(* IEC 61131-3 sources: kauha-loader-autonomy/plc/codesys/src/codesys_only, 3 files *)

(* ---- GVL_IO.st ---- *)
(* Hardware I/O of the 1:8 testbed safety PLC. Map each variable to its channel in
   the device's "I/O Mapping" tab (Raspberry Pi GPIOs device, or the I/O modules of
   your controller). Pin numbers are the testbed wiring in docs/scale/wiring.md.
   Inputs arrive through the 24 V opto-isolated input board (high = 24 V present). *)
VAR_GLOBAL
    (* inputs *)
    xEstopChainOk    : BOOL;   (* IN1  GPIO5:  safety relay K1 contact 33-34, TRUE = chain closed and K1 reset *)
    xRelayFeedbackOk : BOOL;   (* IN2  GPIO6:  K-DRIVE and K-IMPL NC mirror contacts in series, TRUE = both dropped *)
    stScannerIO      : ST_ScannerIO;
                               (* IN3  GPIO12: front_ossd_clear   IN4  GPIO13: rear_ossd_clear
                                  IN5  GPIO19: front_warn_clear   IN6  GPIO20: rear_warn_clear
                                  IN7  GPIO21: side_clear         IN8  GPIO26: under_clear
                                  scanners_ready: IN3..IN8 board "power good" (GPIO4) *)
    (* outputs *)
    xDriveEnable     : BOOL;   (* OUT1 GPIO23: coil of K-DRIVE (motor power and dynamic-brake changeover) *)
    xImplementEnable : BOOL;   (* OUT2 GPIO24: coil of K-IMPL (actuator power) *)
    xFs0, xFs1, xFs2, xFs3, xFs4, xFs5 : BOOL;
                               (* OUT3..OUT8 GPIO16, 17, 22, 27, 18, 14: field-set code bits 0..5 to the
                                  rated scanners' static control inputs (only with USE_SCANNER_IO) *)
    xRunLamp         : BOOL;   (* OUT9 GPIO15: green beacon, machine may move *)
END_VAR

VAR_GLOBAL CONSTANT
    (* FALSE: field bits from the ScannerStatus frame (software evaluator on a hobby lidar, not safety rated).
       TRUE: field bits from rated scanner outputs on stScannerIO. *)
    USE_SCANNER_IO : BOOL := FALSE;
END_VAR

(* ---- FB_CanPort.st ---- *)
(* CAN port for CODESYS Control (Raspberry Pi SL with SocketCAN, or any controller
   with a CAN interface), using the "CAA CAN Low Level" library (namespace CL2).

   Not compiled by the matiec tests: this is the only code that calls a vendor
   library. It moves raw frames between the driver and FB_SafetyNode; every
   check on their content happens in the tested code.

   Library signatures follow the CODESYS online help for CAA CAN Low Level
   3.5.16/3.5.17 (DriverOpenH, CreateMaskReceiver, Read, GetMessageId,
   GetMessageDataPointer, FreeMessage, CreateMessage, Write). If the compiler
   reports a parameter mismatch on another library version, adjust the call here;
   nothing else depends on it. *)

FUNCTION_BLOCK FB_CanPort
VAR_INPUT
    usiNetId   : USINT := 0;       (* CAN interface number: can0 = 0 *)
    uiBaudrate : UINT := 500;      (* kbit/s, as configured on the bus *)
    xReceive   : BOOL;             (* collect the frames waiting in the driver this call *)
    xSend      : BOOL;             (* send tx_id/tx this call *)
    tx_id      : DWORD;
    tx         : ST_Payload;
END_VAR
VAR_OUTPUT
    rx         : ST_RxBatch;       (* frames received since the last call, oldest first *)
    xOpen      : BOOL;
    udiRx      : UDINT;
    udiTx      : UDINT;
    udiErrors  : UDINT;
    udiDropped : UDINT;            (* more than 32 frames waiting in one cycle *)
END_VAR
VAR
    hDriver   : CAA.HANDLE := CAA.gc_hINVALID;
    hReceiver : CAA.HANDLE := CAA.gc_hINVALID;
    hMsg      : CAA.HANDLE;
    eError    : CL2.ERROR;
    ctLeft    : CAA.COUNT;
    pByte     : POINTER TO BYTE;
    i         : INT;
END_VAR

IF hDriver = CAA.gc_hINVALID THEN
    hDriver := CL2.DriverOpenH(usiNetId := usiNetId, uiBaudrate := uiBaudrate, xSupport29Bits := TRUE,
                               ctMessages := 64, peError := ADR(eError));
    IF hDriver <> CAA.gc_hINVALID THEN
        (* every extended-ID data frame that this node did not send itself *)
        hReceiver := CL2.CreateMaskReceiver(hDriver := hDriver,
                                            cobIdValue := 0, cobIdMask := 0,
                                            xRTRValue := FALSE, xRTRMask := TRUE,
                                            x29BitIdValue := TRUE, x29BitIdMask := TRUE,
                                            xTransmitValue := FALSE, xTransmitMask := TRUE,
                                            xAlwaysNewest := FALSE, eEvent := CB.EVENT.NO_EVENT,
                                            xEnableSyncWindow := FALSE, peError := ADR(eError));
    END_IF
END_IF
xOpen := (hDriver <> CAA.gc_hINVALID) AND (hReceiver <> CAA.gc_hINVALID);

IF xReceive THEN
    rx.n := 0;
END_IF
WHILE xOpen AND xReceive DO
    hMsg := CL2.Read(hReceiverId := hReceiver, pctMsgLeft := ADR(ctLeft), peError := ADR(eError));
    IF hMsg = CAA.gc_hINVALID THEN
        EXIT;
    END_IF
    IF rx.n < 32 THEN
        rx.f[rx.n].id := CL2.GetMessageId(hMessage := hMsg, peError := ADR(eError));
        pByte := CL2.GetMessageDataPointer(hMessage := hMsg, peError := ADR(eError));
        FOR i := 0 TO 7 DO
            rx.f[rx.n].data.b[i] := (pByte + i)^;
        END_FOR
        rx.n := rx.n + 1;
        udiRx := udiRx + 1;
    ELSE
        udiDropped := udiDropped + 1;   (* dropped frames read as missing: the E2E checks see them as lost *)
    END_IF
    CL2.FreeMessage(hMessage := hMsg, peError := ADR(eError));
END_WHILE

IF xSend AND xOpen THEN
    hMsg := CL2.CreateMessage(hDriver := hDriver, cobID := tx_id, usiLength := 8, xRTR := FALSE,
                              x29BitID := TRUE, peError := ADR(eError));
    IF hMsg <> CAA.gc_hINVALID THEN
        pByte := CL2.GetMessageDataPointer(hMessage := hMsg, peError := ADR(eError));
        FOR i := 0 TO 7 DO
            (pByte + i)^ := tx.b[i];
        END_FOR
        eError := CL2.Write(hDriver := hDriver, hMessage := hMsg, usiPriority := 0, xEnableSyncWindow := FALSE);
        IF eError = CL2.ERROR.NO_ERROR THEN
            udiTx := udiTx + 1;
        ELSE
            udiErrors := udiErrors + 1;
        END_IF
    ELSE
        udiErrors := udiErrors + 1;
    END_IF
END_IF
END_FUNCTION_BLOCK

(* ---- PRG_Main.st ---- *)
(* Main program of the testbed safety PLC. Run it in a cyclic task of 25 ms
   (Task configuration: "SafetyTask", cyclic, t#25ms, priority 1, watchdog 50 ms).

   Choose the configuration list for the profile that matches the hardware:
     CFG_SCALE8_EVALUATOR  hobby lidar + software field evaluator (first tests)
     CFG_SCALE8_NANOSCAN3  rated SICK nanoScan3 I/O scanners (set USE_SCANNER_IO := TRUE)
     CFG_FULL              the full-size machine (reference only)
   The profiles are generated by `python -m kauha.scale.profile` from the same
   numbers the twin and the proofs use. *)

PROGRAM PRG_Main
VAR
    can  : FB_CanPort;
    node : FB_SafetyNode;
    t    : LREAL;
    relayCheck : TON;          (* a stop must be followed by both relays dropping *)
    xRelayFault : BOOL;
END_VAR

t := TIME_TO_LREAL(TIME()) / 1000.0;

can(xReceive := TRUE, xSend := FALSE);

node(cfg := CFG_SCALE8_EVALUATOR,
     t := t,
     rx := can.rx,
     estop_chain_ok := GVL_IO.xEstopChainOk AND NOT xRelayFault,
     use_scanner_io := GVL_IO.USE_SCANNER_IO,
     scanner_io := GVL_IO.stScannerIO);

GVL_IO.xDriveEnable := node.drive_enable;
GVL_IO.xImplementEnable := node.implement_enable;
GVL_IO.xRunLamp := node.drive_enable;
GVL_IO.xFs0 := (node.field_set_code AND 16#01) <> 0;
GVL_IO.xFs1 := (node.field_set_code AND 16#02) <> 0;
GVL_IO.xFs2 := (node.field_set_code AND 16#04) <> 0;
GVL_IO.xFs3 := (node.field_set_code AND 16#08) <> 0;
GVL_IO.xFs4 := (node.field_set_code AND 16#10) <> 0;
GVL_IO.xFs5 := (node.field_set_code AND 16#20) <> 0;

(* Relay monitoring: with both coils off, the mirror contacts must close within 100 ms.
   A welded contact latches a fault that reads as an e-stop until power cycle. *)
relayCheck(IN := NOT GVL_IO.xDriveEnable AND NOT GVL_IO.xImplementEnable AND NOT GVL_IO.xRelayFeedbackOk,
           PT := T#100MS);
IF relayCheck.Q THEN
    xRelayFault := TRUE;
END_IF

can(xReceive := FALSE, xSend := TRUE, tx_id := node.tx_id, tx := node.tx);
END_PROGRAM
